// TIA Portal project "Three_Pump_Booster_Control" (V19)
// Three-pump VFD booster station with PID pressure control, lead/lag sequencing and WinCC HMI

(* hardware
DEVICE "S7-1500/ET200MP station_1"  S7-1500 station
   slot 0: "Rail_0"  Rack  6ES7 590-1***0-0AA0
   slot 1: "PLC_Booster"  CPU 1511-1 PN  6ES7 511-1AK02-0AB0  V2.9
      slot 3: "CPU display_1"  6ES7591-1AA00-0AA0
      slot 32768: "PROFINET interface_1"  X1
         slot 32769: "Port_1"  X1 P1
         slot 32770: "Port_2"  X1 P2
      slot 34817: "Virtual CP interface port_1"  Virtual CP interface port  Virtual CP interface port
DEVICE "HMI_Booster"  SIMATIC PC station
   slot 0: "SIMATIC PC station"  Rail  SIMATIC PC-Station  V1.0
      slot 125: "Stationmanager"  Station_Manager  V6.0.4
   slot 1: "HMI_RT_1"  WinCC RT Advanced  6AV2 104-0xxxx-xxxx  17.0.0.0
      slot 33792: "Computer interface"  Host interface
   slot 2: "IE general_1"  IE General  IE_CP  V8.2.0
      slot 1: "PROFINET interface"  IEGeneral.Interface.8.2.0
*)

// ===== PLC "PLC_Booster"  CPU 1511-1 PN =====

TYPE "UDT_Pump"
   STRUCT
      CmdRun : Bool;
      CmdSpeedPct : Real;
      FbRunning : Bool;
      FbFault : Bool;
      FbSpeedPct : Real;
      RunHours : Real;
      Role : Int;
   END_STRUCT;
END_TYPE

DATA_BLOCK "DB_Pumps"   // DB1
{ S7_Optimized_Access := 'TRUE' }
VERSION : 0.1
   VAR
      Pump1 : "UDT_Pump";
      Pump2 : "UDT_Pump";
      Pump3 : "UDT_Pump";
   END_VAR
BEGIN
END_DATA_BLOCK

DATA_BLOCK "DB_System"   // DB2
{ S7_Optimized_Access := 'TRUE' }
VERSION : 0.1
   VAR
      SystemRun : Bool;
      AutoMode : Bool := TRUE;
      SimEnable : Bool := TRUE;
      PressureSP : Real := 4.0;
      PressurePV : Real;
      PIDOutputPct : Real;
      DemandPct : Real := 35.0;
      PressureHighSP : Real := 6.0;
      PressureLowSP : Real := 2.0;
      PIDMode : Int := 4;
      PIDModeActivate : Bool;
      Pump1RunReq : Bool;
      Pump2RunReq : Bool;
      Pump3RunReq : Bool;
      Pump1SpeedReq : Real;
      Pump2SpeedReq : Real;
      Pump3SpeedReq : Real;
      PumpPermissive : Bool := TRUE;
      Pump1FaultAlarm : Bool;
      Pump2FaultAlarm : Bool;
      Pump3FaultAlarm : Bool;
      PressureHighAlarm : Bool;
      PressureLowAlarm : Bool;
      AnyAlarm : Bool;
      Pump1Role : Int;
      Pump2Role : Int;
      Pump3Role : Int;
      AlarmWord : Word := W#16#0000;
   END_VAR
BEGIN
END_DATA_BLOCK

DATA_BLOCK "DB_Pump1_Control"   // DB3
{ S7_Optimized_Access := 'TRUE' }
VERSION : 0.1
// stored: InstanceOfName FB_PumpControl
"FB_PumpControl"
BEGIN
END_DATA_BLOCK

DATA_BLOCK "DB_Pump2_Control"   // DB4
{ S7_Optimized_Access := 'TRUE' }
VERSION : 0.1
// stored: InstanceOfName FB_PumpControl
"FB_PumpControl"
BEGIN
END_DATA_BLOCK

DATA_BLOCK "DB_Pump3_Control"   // DB5
{ S7_Optimized_Access := 'TRUE' }
VERSION : 0.1
// stored: InstanceOfName FB_PumpControl
"FB_PumpControl"
BEGIN
END_DATA_BLOCK

DATA_BLOCK "DB_ProcessSimulation"   // DB6
{ S7_Optimized_Access := 'TRUE' }
VERSION : 0.1
// stored: InstanceOfName FB_ProcessSimulation
"FB_ProcessSimulation"
BEGIN
END_DATA_BLOCK

DATA_BLOCK "DB_PumpManager"   // DB8
{ S7_Optimized_Access := 'TRUE' }
VERSION : 0.1
// stored: InstanceOfName FB_PumpManager
"FB_PumpManager"
BEGIN
END_DATA_BLOCK

DATA_BLOCK "DB_AlarmManager"   // DB9
{ S7_Optimized_Access := 'TRUE' }
VERSION : 0.1
// stored: InstanceOfName FB_AlarmManager
"FB_AlarmManager"
BEGIN
END_DATA_BLOCK

FUNCTION_BLOCK "FB_PumpControl"   // FB1, LAD
{ S7_Optimized_Access := 'TRUE' }
VERSION : 0.1
   VAR_INPUT
      RunRequest : Bool;
      SpeedRequestPct : Real;
      Permissive : Bool;
   END_VAR
   VAR_IN_OUT
      Pump : "UDT_Pump";
   END_VAR
   VAR_TEMP
      LimitedSpeedPct : Real;
   END_VAR
BEGIN

REGION Network 1: VFD Run Command
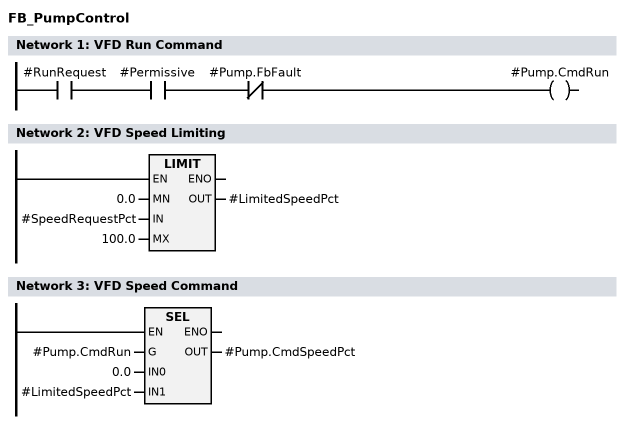
   RUNG wire#powerrail
      Contact( #RunRequest )
      Contact( #Permissive )
      I_Contact( #Pump.FbFault )
      Coil( #Pump.CmdRun )
   END_RUNG
   // the same network as SCL:
   #Pump.CmdRun := #RunRequest AND #Permissive AND NOT #Pump.FbFault;
END_REGION

REGION Network 2: VFD Speed Limiting
   #LimitedSpeedPct := LIMIT(MN := 0.0, IN := #SpeedRequestPct, MX := 100.0);
END_REGION

REGION Network 3: VFD Speed Command
   #Pump.CmdSpeedPct := SEL(G := #Pump.CmdRun, IN0 := 0.0, IN1 := #LimitedSpeedPct);
END_REGION
END_FUNCTION_BLOCK

FUNCTION_BLOCK "FB_ProcessSimulation"   // FB2, SCL
{ S7_Optimized_Access := 'TRUE' }
VERSION : 0.1
   VAR_INPUT
      SimEnable : Bool;
      DemandPct : Real;
   END_VAR
   VAR_IN_OUT
      Pump1 : "UDT_Pump";
      Pump2 : "UDT_Pump";
      Pump3 : "UDT_Pump";
      PressurePV : Real;
   END_VAR
   VAR_TEMP
      TargetSpeed1 : Real;
      TargetSpeed2 : Real;
      TargetSpeed3 : Real;
      TotalFlow : Real;
      DemandLimited : Real;
   END_VAR
BEGIN

   IF NOT #SimEnable THEN
       // Reset simulated process
       #Pump1.FbSpeedPct := 0.0;
       #Pump2.FbSpeedPct := 0.0;
       #Pump3.FbSpeedPct := 0.0;

       #Pump1.FbRunning := FALSE;
       #Pump2.FbRunning := FALSE;
       #Pump3.FbRunning := FALSE;

       #PressurePV := 0.0;

   ELSE
       // Determine requested VFD speeds
       #TargetSpeed1 := 0.0;
       #TargetSpeed2 := 0.0;
       #TargetSpeed3 := 0.0;

       IF #Pump1.CmdRun AND NOT #Pump1.FbFault THEN
           #TargetSpeed1 := #Pump1.CmdSpeedPct;
       END_IF;

       IF #Pump2.CmdRun AND NOT #Pump2.FbFault THEN
           #TargetSpeed2 := #Pump2.CmdSpeedPct;
       END_IF;

       IF #Pump3.CmdRun AND NOT #Pump3.FbFault THEN
           #TargetSpeed3 := #Pump3.CmdSpeedPct;
       END_IF;

       // Simulate VFD acceleration and deceleration
       #Pump1.FbSpeedPct := #Pump1.FbSpeedPct +
       0.2 * (#TargetSpeed1 - #Pump1.FbSpeedPct);

       #Pump2.FbSpeedPct := #Pump2.FbSpeedPct +
       0.2 * (#TargetSpeed2 - #Pump2.FbSpeedPct);

       #Pump3.FbSpeedPct := #Pump3.FbSpeedPct +
       0.2 * (#TargetSpeed3 - #Pump3.FbSpeedPct);

       // Simulated running feedback
       #Pump1.FbRunning := #Pump1.FbSpeedPct > 1.0;
       #Pump2.FbRunning := #Pump2.FbSpeedPct > 1.0;
       #Pump3.FbRunning := #Pump3.FbSpeedPct > 1.0;

       // Combined pump flow (arbitrary simulation units)
       #TotalFlow := 1.1 * (
       #Pump1.FbSpeedPct +
       #Pump2.FbSpeedPct +
       #Pump3.FbSpeedPct
       );

       // Limit simulated water demand
       #DemandLimited := #DemandPct;

       IF #DemandLimited < 0.0 THEN
           #DemandLimited := 0.0;
       ELSIF #DemandLimited > 100.0 THEN
           #DemandLimited := 100.0;
       END_IF;

       // Pressure model: designed for a 100 ms cycle
       #PressurePV := #PressurePV + 0.004 *
       (#TotalFlow - #DemandLimited -
       12.0 * #PressurePV);

       // Limit simulated pressure to 0-10 bar
       IF #PressurePV < 0.0 THEN
           #PressurePV := 0.0;
       ELSIF #PressurePV > 10.0 THEN
           #PressurePV := 10.0;
       END_IF;

   END_IF;
END_FUNCTION_BLOCK

FUNCTION_BLOCK "FB_PumpManager"   // FB3, SCL
{ S7_Optimized_Access := 'TRUE' }
VERSION : 0.1
   VAR_INPUT
      SystemRun : Bool;
      AutoMode : Bool;
      SimEnable : Bool;
      PumpPermissive : Bool;
      PressureSP : Real;
      PressurePV : Real;
      PIDOutputPct : Real;
      Pump1Fault : Bool;
      Pump2Fault : Bool;
      Pump3Fault : Bool;
   END_VAR
   VAR_OUTPUT
      Pump1RunReq : Bool;
      Pump2RunReq : Bool;
      Pump3RunReq : Bool;
      Pump1SpeedReq : Real;
      Pump2SpeedReq : Real;
      Pump3SpeedReq : Real;
      Pump1Role : Int;
      Pump2Role : Int;
      Pump3Role : Int;
   END_VAR
   VAR
      LagActive : Bool;
      StageUpCount : Int := 0;
      StageDownCount : Int;
      LeadPumpNo : Int := 1;
      LagPumpNo : Int;
   END_VAR
   VAR_TEMP
      PreviousLead : Int;
   END_VAR
BEGIN

   (* Default pump commands *)
   #Pump1RunReq := FALSE;
   #Pump2RunReq := FALSE;
   #Pump3RunReq := FALSE;

   #Pump1SpeedReq := 0.0;
   #Pump2SpeedReq := 0.0;
   #Pump3SpeedReq := 0.0;

   IF NOT (#SystemRun AND #AutoMode AND
       #SimEnable AND #PumpPermissive) THEN

       // Reset assignments when system stops
       #LeadPumpNo := 1;
       #LagPumpNo := 0;
       #LagActive := FALSE;
       #StageUpCount := 0;
       #StageDownCount := 0;

   ELSE

       #PreviousLead := #LeadPumpNo;

       // Check the selected lead pump
       CASE #LeadPumpNo OF

           1:
               IF #Pump1Fault THEN
                   IF NOT #Pump3Fault THEN
                       #LeadPumpNo := 3;
                   ELSIF NOT #Pump2Fault THEN
                       #LeadPumpNo := 2;
                   ELSE
                       #LeadPumpNo := 0;
                   END_IF;
               END_IF;

           2:
               IF #Pump2Fault THEN
                   IF NOT #Pump3Fault THEN
                       #LeadPumpNo := 3;
                   ELSIF NOT #Pump1Fault THEN
                       #LeadPumpNo := 1;
                   ELSE
                       #LeadPumpNo := 0;
                   END_IF;
               END_IF;

           3:
               IF #Pump3Fault THEN
                   IF NOT #Pump2Fault THEN
                       #LeadPumpNo := 2;
                   ELSIF NOT #Pump1Fault THEN
                       #LeadPumpNo := 1;
                   ELSE
                       #LeadPumpNo := 0;
                   END_IF;
               END_IF;

           ELSE
               // Recover when a pump becomes available
               IF NOT #Pump1Fault THEN
                   #LeadPumpNo := 1;
               ELSIF NOT #Pump3Fault THEN
                   #LeadPumpNo := 3;
               ELSIF NOT #Pump2Fault THEN
                   #LeadPumpNo := 2;
               ELSE
                   #LeadPumpNo := 0;
               END_IF;

       END_CASE;

       // Reset staging after lead changeover
       IF #LeadPumpNo <> #PreviousLead THEN
           #LagActive := FALSE;
           #LagPumpNo := 0;
           #StageUpCount := 0;
           #StageDownCount := 0;
       END_IF;

       // Check an active assist pump for faults
       IF #LagActive THEN

           IF ((#LagPumpNo = 1) AND #Pump1Fault) OR
               ((#LagPumpNo = 2) AND #Pump2Fault) OR
               ((#LagPumpNo = 3) AND #Pump3Fault) OR
               (#LagPumpNo = #LeadPumpNo) THEN

               #LagPumpNo := 0;

               // Select another healthy assist pump
               CASE #LeadPumpNo OF

                   1:
                       IF NOT #Pump2Fault THEN
                           #LagPumpNo := 2;
                       ELSIF NOT #Pump3Fault THEN
                           #LagPumpNo := 3;
                       END_IF;

                   2:
                       IF NOT #Pump3Fault THEN
                           #LagPumpNo := 3;
                       ELSIF NOT #Pump1Fault THEN
                           #LagPumpNo := 1;
                       END_IF;

                   3:
                       IF NOT #Pump2Fault THEN
                           #LagPumpNo := 2;
                       ELSIF NOT #Pump1Fault THEN
                           #LagPumpNo := 1;
                       END_IF;

               END_CASE;

               IF #LagPumpNo = 0 THEN
                   #LagActive := FALSE;
               END_IF;

           END_IF;

       END_IF;

       // Automatic lag pump staging
       IF NOT #LagActive THEN

           #StageDownCount := 0;

           IF (#LeadPumpNo <> 0) AND
               (#PIDOutputPct >= 95.0) AND
               (#PressurePV < (#PressureSP - 0.2)) THEN

               IF #StageUpCount < 50 THEN
                   #StageUpCount := #StageUpCount + 1;
               END_IF;

           ELSE
               #StageUpCount := 0;
           END_IF;

           IF #StageUpCount >= 50 THEN

               #LagPumpNo := 0;

               CASE #LeadPumpNo OF

                   1:
                       IF NOT #Pump2Fault THEN
                           #LagPumpNo := 2;
                       ELSIF NOT #Pump3Fault THEN
                           #LagPumpNo := 3;
                       END_IF;

                   2:
                       IF NOT #Pump3Fault THEN
                           #LagPumpNo := 3;
                       ELSIF NOT #Pump1Fault THEN
                           #LagPumpNo := 1;
                       END_IF;

                   3:
                       IF NOT #Pump2Fault THEN
                           #LagPumpNo := 2;
                       ELSIF NOT #Pump1Fault THEN
                           #LagPumpNo := 1;
                       END_IF;

               END_CASE;

               #LagActive := (#LagPumpNo <> 0);
               #StageUpCount := 0;

           END_IF;

       ELSE

           #StageUpCount := 0;

           IF (#PIDOutputPct <= 50.0) AND
               (#PressurePV >= (#PressureSP - 0.1)) THEN

               IF #StageDownCount < 100 THEN
                   #StageDownCount := #StageDownCount + 1;
               END_IF;

           ELSE
               #StageDownCount := 0;
           END_IF;

           IF #StageDownCount >= 100 THEN
               #LagActive := FALSE;
               #LagPumpNo := 0;
               #StageDownCount := 0;
           END_IF;

       END_IF;

       // Assign PID speed to selected lead pump
       CASE #LeadPumpNo OF

           1:
               #Pump1RunReq := TRUE;
               #Pump1SpeedReq := #PIDOutputPct;

           2:
               #Pump2RunReq := TRUE;
               #Pump2SpeedReq := #PIDOutputPct;

           3:
               #Pump3RunReq := TRUE;
               #Pump3SpeedReq := #PIDOutputPct;

       END_CASE;

       // Assign fixed 30% speed to assist pump
       IF #LagActive THEN

           CASE #LagPumpNo OF

               1:
                   #Pump1RunReq := TRUE;
                   #Pump1SpeedReq := 30.0;

               2:
                   #Pump2RunReq := TRUE;
                   #Pump2SpeedReq := 30.0;

               3:
                   #Pump3RunReq := TRUE;
                   #Pump3SpeedReq := 30.0;

           END_CASE;

       END_IF;

   END_IF;


   // Default: All pumps on standby
   #Pump1Role := 0;
   #Pump2Role := 0;
   #Pump3Role := 0;

   // Assign operating roles when system enabled
   IF #SystemRun AND #AutoMode AND
       #SimEnable AND #PumpPermissive THEN

       // Lead pump role
       CASE #LeadPumpNo OF
           1:
               #Pump1Role := 1;
           2:
               #Pump2Role := 1;
           3:
               #Pump3Role := 1;
       END_CASE;

       // Assist pump role
       IF #LagActive THEN
           CASE #LagPumpNo OF
               1:
                   #Pump1Role := 2;
               2:
                   #Pump2Role := 2;
               3:
                   #Pump3Role := 2;
           END_CASE;
       END_IF;

   END_IF;

   // Fault indication takes priority
   IF #Pump1Fault THEN
       #Pump1Role := 3;
   END_IF;

   IF #Pump2Fault THEN
       #Pump2Role := 3;
   END_IF;

   IF #Pump3Fault THEN
       #Pump3Role := 3;
   END_IF;
END_FUNCTION_BLOCK

FUNCTION_BLOCK "FB_AlarmManager"   // FB4, SCL
{ S7_Optimized_Access := 'TRUE' }
VERSION : 0.1
   VAR_INPUT
      SystemRun : Bool;
      PressurePV : Real;
      PressureHighSP : Real;
      PressureLowSP : Real;
      Pump1Fault : Bool;
      Pump2Fault : Bool;
      Pump3Fault : Bool;
   END_VAR
   VAR_OUTPUT
      Pump1FaultAlarm : Bool;
      Pump2FaultAlarm : Bool;
      Pump3FaultAlarm : Bool;
      PressureHighAlarm : Bool;
      PressureLowAlarm : Bool;
      AnyAlarm : Bool;
      AlarmWord : Word;
   END_VAR
   VAR
      LowPressureCount : Int;
   END_VAR
BEGIN

   // Individual pump fault alarms
   #Pump1FaultAlarm := #Pump1Fault;
   #Pump2FaultAlarm := #Pump2Fault;
   #Pump3FaultAlarm := #Pump3Fault;

   // High pressure alarm with hysteresis
   IF #PressurePV >= #PressureHighSP THEN
       #PressureHighAlarm := TRUE;
   ELSIF #PressurePV <= (#PressureHighSP - 0.2) THEN
       #PressureHighAlarm := FALSE;
   END_IF;

   // Low pressure alarm with 10-second delay
   // FB must execute every 100 ms
   IF NOT #SystemRun THEN
       #LowPressureCount := 0;
       #PressureLowAlarm := FALSE;

   ELSIF #PressurePV < #PressureLowSP THEN
       IF #LowPressureCount < 100 THEN
           #LowPressureCount := #LowPressureCount + 1;
       END_IF;

       IF #LowPressureCount >= 100 THEN
           #PressureLowAlarm := TRUE;
       END_IF;

   ELSE
       #LowPressureCount := 0;

       IF #PressurePV >= (#PressureLowSP + 0.2) THEN
           #PressureLowAlarm := FALSE;
       END_IF;
   END_IF;

   // General alarm indication
   #AnyAlarm :=
   #Pump1FaultAlarm OR
   #Pump2FaultAlarm OR
   #Pump3FaultAlarm OR
   #PressureHighAlarm OR
   #PressureLowAlarm;



   // Pack individual alarm signals
   // into one WinCC alarm trigger word

   #AlarmWord := W#16#0000;

   IF #Pump1FaultAlarm THEN
       #AlarmWord := #AlarmWord OR W#16#0001;
   END_IF;

   IF #Pump2FaultAlarm THEN
       #AlarmWord := #AlarmWord OR W#16#0002;
   END_IF;

   IF #Pump3FaultAlarm THEN
       #AlarmWord := #AlarmWord OR W#16#0004;
   END_IF;

   IF #PressureHighAlarm THEN
       #AlarmWord := #AlarmWord OR W#16#0008;
   END_IF;

   IF #PressureLowAlarm THEN
       #AlarmWord := #AlarmWord OR W#16#0010;
   END_IF;
END_FUNCTION_BLOCK

ORGANIZATION_BLOCK "Main"   // OB1, LAD, ProgramCycle
TITLE = "Main Program Sweep (Cycle)"
{ S7_Optimized_Access := 'TRUE' }
VERSION : 0.1
   VAR_INPUT
      Initial_Call : Bool;   // Initial call of this OB
      Remanence : Bool;   // =True, if remanent data are available
   END_VAR
BEGIN

REGION Network 1: Pump 1 VFD Control
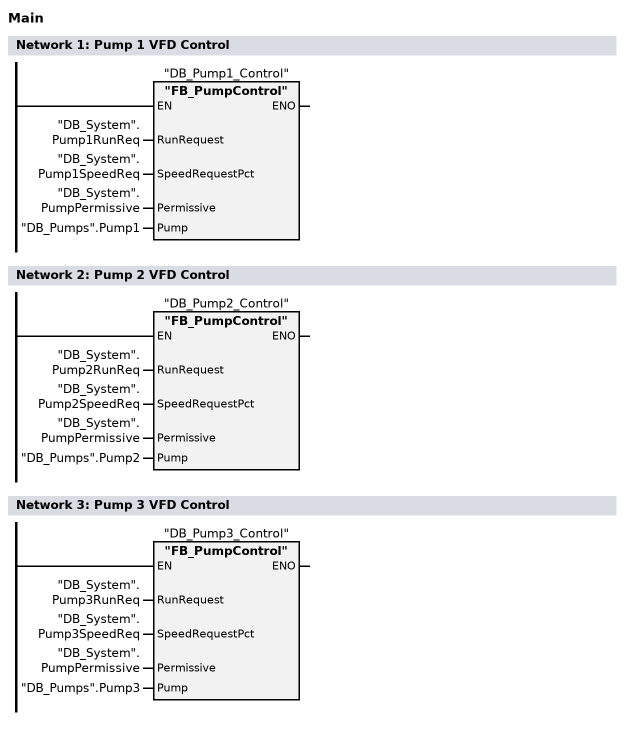
   RUNG wire#powerrail
      "DB_Pump1_Control"(RunRequest := "DB_System".Pump1RunReq, SpeedRequestPct := "DB_System".Pump1SpeedReq, Permissive := "DB_System".PumpPermissive, Pump := "DB_Pumps".Pump1)
   END_RUNG
   // the same network as SCL:
   "DB_Pump1_Control"(RunRequest := "DB_System".Pump1RunReq,   // "FB_PumpControl"
                      SpeedRequestPct := "DB_System".Pump1SpeedReq,
                      Permissive := "DB_System".PumpPermissive,
                      Pump := "DB_Pumps".Pump1);
END_REGION

REGION Network 2: Pump 2 VFD Control
   RUNG wire#powerrail
      "DB_Pump2_Control"(RunRequest := "DB_System".Pump2RunReq, SpeedRequestPct := "DB_System".Pump2SpeedReq, Permissive := "DB_System".PumpPermissive, Pump := "DB_Pumps".Pump2)
   END_RUNG
   // the same network as SCL:
   "DB_Pump2_Control"(RunRequest := "DB_System".Pump2RunReq,   // "FB_PumpControl"
                      SpeedRequestPct := "DB_System".Pump2SpeedReq,
                      Permissive := "DB_System".PumpPermissive,
                      Pump := "DB_Pumps".Pump2);
END_REGION

REGION Network 3: Pump 3 VFD Control
   RUNG wire#powerrail
      "DB_Pump3_Control"(RunRequest := "DB_System".Pump3RunReq, SpeedRequestPct := "DB_System".Pump3SpeedReq, Permissive := "DB_System".PumpPermissive, Pump := "DB_Pumps".Pump3)
   END_RUNG
   // the same network as SCL:
   "DB_Pump3_Control"(RunRequest := "DB_System".Pump3RunReq,   // "FB_PumpControl"
                      SpeedRequestPct := "DB_System".Pump3SpeedReq,
                      Permissive := "DB_System".PumpPermissive,
                      Pump := "DB_Pumps".Pump3);
END_REGION
END_ORGANIZATION_BLOCK

ORGANIZATION_BLOCK "OB30_ProcessControl"   // OB30, LAD, CyclicInterrupt
{ S7_Optimized_Access := 'TRUE' }
VERSION : 0.1
   VAR_INPUT
      Initial_Call : Bool;   // Initial call of this OB
      Event_Count : Int;   // Events discarded
   END_VAR
BEGIN

REGION Network 1: Hydraulic Process Simulation
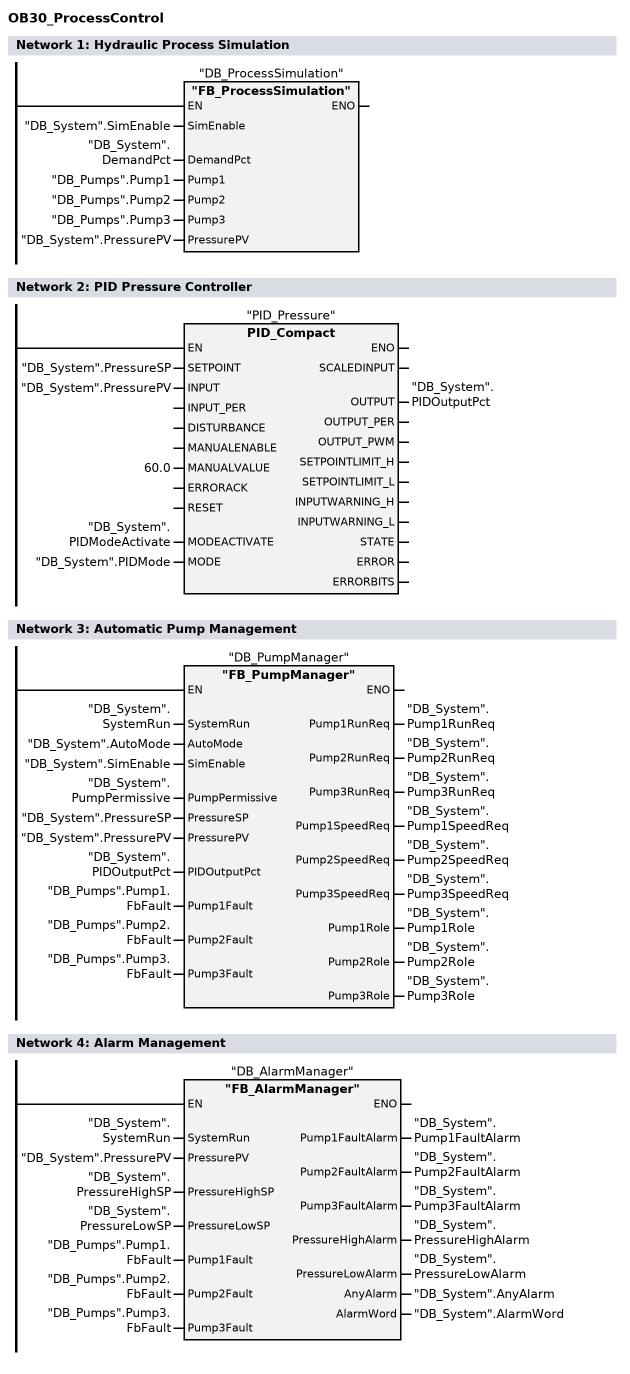
   RUNG wire#powerrail
      "DB_ProcessSimulation"(SimEnable := "DB_System".SimEnable, DemandPct := "DB_System".DemandPct, Pump1 := "DB_Pumps".Pump1, Pump2 := "DB_Pumps".Pump2, Pump3 := "DB_Pumps".Pump3, PressurePV := "DB_System".PressurePV)
   END_RUNG
   // the same network as SCL:
   "DB_ProcessSimulation"(SimEnable := "DB_System".SimEnable,   // "FB_ProcessSimulation"
                          DemandPct := "DB_System".DemandPct,
                          Pump1 := "DB_Pumps".Pump1,
                          Pump2 := "DB_Pumps".Pump2,
                          Pump3 := "DB_Pumps".Pump3,
                          PressurePV := "DB_System".PressurePV);
END_REGION

REGION Network 2: PID Pressure Controller
   "PID_Pressure"(Setpoint := "DB_System".PressureSP,   // PID_Compact
                  Input := "DB_System".PressurePV,
                  ManualValue := 60.0,
                  ModeActivate := "DB_System".PIDModeActivate,
                  Mode := "DB_System".PIDMode,
                  Output => "DB_System".PIDOutputPct);
END_REGION

REGION Network 3: Automatic Pump Management
   RUNG wire#powerrail
      "DB_PumpManager"(SystemRun := "DB_System".SystemRun, AutoMode := "DB_System".AutoMode, SimEnable := "DB_System".SimEnable, PumpPermissive := "DB_System".PumpPermissive, PressureSP := "DB_System".PressureSP, PressurePV := "DB_System".PressurePV, PIDOutputPct := "DB_System".PIDOutputPct, Pump1Fault := "DB_Pumps".Pump1.FbFault, Pump2Fault := "DB_Pumps".Pump2.FbFault, Pump3Fault := "DB_Pumps".Pump3.FbFault, Pump1RunReq => "DB_System".Pump1RunReq, Pump2RunReq => "DB_System".Pump2RunReq, Pump3RunReq => "DB_System".Pump3RunReq, Pump1SpeedReq => "DB_System".Pump1SpeedReq, Pump2SpeedReq => "DB_System".Pump2SpeedReq, Pump3SpeedReq => "DB_System".Pump3SpeedReq, Pump1Role => "DB_System".Pump1Role, Pump2Role => "DB_System".Pump2Role, Pump3Role => "DB_System".Pump3Role)
   END_RUNG
   // the same network as SCL:
   "DB_PumpManager"(SystemRun := "DB_System".SystemRun,   // "FB_PumpManager"
                    AutoMode := "DB_System".AutoMode,
                    SimEnable := "DB_System".SimEnable,
                    PumpPermissive := "DB_System".PumpPermissive,
                    PressureSP := "DB_System".PressureSP,
                    PressurePV := "DB_System".PressurePV,
                    PIDOutputPct := "DB_System".PIDOutputPct,
                    Pump1Fault := "DB_Pumps".Pump1.FbFault,
                    Pump2Fault := "DB_Pumps".Pump2.FbFault,
                    Pump3Fault := "DB_Pumps".Pump3.FbFault,
                    Pump1RunReq => "DB_System".Pump1RunReq,
                    Pump2RunReq => "DB_System".Pump2RunReq,
                    Pump3RunReq => "DB_System".Pump3RunReq,
                    Pump1SpeedReq => "DB_System".Pump1SpeedReq,
                    Pump2SpeedReq => "DB_System".Pump2SpeedReq,
                    Pump3SpeedReq => "DB_System".Pump3SpeedReq,
                    Pump1Role => "DB_System".Pump1Role,
                    Pump2Role => "DB_System".Pump2Role,
                    Pump3Role => "DB_System".Pump3Role);
END_REGION

REGION Network 4: Alarm Management
   RUNG wire#powerrail
      "DB_AlarmManager"(SystemRun := "DB_System".SystemRun, PressurePV := "DB_System".PressurePV, PressureHighSP := "DB_System".PressureHighSP, PressureLowSP := "DB_System".PressureLowSP, Pump1Fault := "DB_Pumps".Pump1.FbFault, Pump2Fault := "DB_Pumps".Pump2.FbFault, Pump3Fault := "DB_Pumps".Pump3.FbFault, Pump1FaultAlarm => "DB_System".Pump1FaultAlarm, Pump2FaultAlarm => "DB_System".Pump2FaultAlarm, Pump3FaultAlarm => "DB_System".Pump3FaultAlarm, PressureHighAlarm => "DB_System".PressureHighAlarm, PressureLowAlarm => "DB_System".PressureLowAlarm, AnyAlarm => "DB_System".AnyAlarm, AlarmWord => "DB_System".AlarmWord)
   END_RUNG
   // the same network as SCL:
   "DB_AlarmManager"(SystemRun := "DB_System".SystemRun,   // "FB_AlarmManager"
                     PressurePV := "DB_System".PressurePV,
                     PressureHighSP := "DB_System".PressureHighSP,
                     PressureLowSP := "DB_System".PressureLowSP,
                     Pump1Fault := "DB_Pumps".Pump1.FbFault,
                     Pump2Fault := "DB_Pumps".Pump2.FbFault,
                     Pump3Fault := "DB_Pumps".Pump3.FbFault,
                     Pump1FaultAlarm => "DB_System".Pump1FaultAlarm,
                     Pump2FaultAlarm => "DB_System".Pump2FaultAlarm,
                     Pump3FaultAlarm => "DB_System".Pump3FaultAlarm,
                     PressureHighAlarm => "DB_System".PressureHighAlarm,
                     PressureLowAlarm => "DB_System".PressureLowAlarm,
                     AnyAlarm => "DB_System".AnyAlarm,
                     AlarmWord => "DB_System".AlarmWord);
END_REGION
END_ORGANIZATION_BLOCK

(* ===== HMI "HMI_RT_1" =====
system functions are stored by id; their names below are inferred from use
connection "HMI_Connection_1": ETHERNET, S7_1500_OMS

HMI tags "Default tag table"
   "HMI_PressurePV" : Real = PLC DB_System.PressurePV AT %DB1.DBD0, 1 s
   "HMI_PressureSP" : Real = PLC DB_System.PressureSP AT %DB1.DBD0, 1 s
   "HMI_TestValue" : Real AT %DB1.DBD0
   "HMI_P1_Running" : Bool = PLC DB_Pumps.Pump1.FbRunning AT %DB1.DBX0.0, 1 s
   "HMI_P2_Running" : Bool = PLC DB_Pumps.Pump2.FbRunning AT %DB1.DBX0.0, 1 s
   "HMI_P3_Running" : Bool = PLC DB_Pumps.Pump3.FbRunning AT %DB1.DBX0.0, 1 s
   "HMI_P1_Speed" : Real = PLC DB_Pumps.Pump1.FbSpeedPct AT %DB1.DBX0.0, 1 s
   "HMI_P2_Speed" : Real = PLC DB_Pumps.Pump2.FbSpeedPct AT %DB1.DBD0, 1 s
   "HMI_P3_Speed" : Real = PLC DB_Pumps.Pump3.FbSpeedPct AT %DB1.DBD0, 1 s
   "HMI_SystemRun" : Bool = PLC DB_System.SystemRun AT %DB1.DBX0.0, 1 s
   "HMI_PIDOutput" : Real = PLC DB_System.PIDOutputPct AT %DB1.DBD0, 1 s
   "HMI_P1_Role" : Int = PLC DB_System.Pump1Role AT %DB1.DBW0, 1 s
   "HMI_P2_Role" : Int = PLC DB_System.Pump2Role AT %DB1.DBW0, 1 s
   "HMI_P3_Role" : Int = PLC DB_System.Pump3Role AT %DB1.DBW0, 1 s
   "HMI_DemandPct" : Real = PLC DB_System.DemandPct AT %DB1.DBD0, 1 s
   "HMI_AutoMode" : Bool = PLC DB_System.AutoMode AT %DB1.DBX0.0, 1 s
   "HMI_AnyAlarm" : Bool = PLC DB_System.AnyAlarm AT %DB1.DBX0.0, 1 s
   "PID_ACTIVE" : Bool = PLC DB_System.PIDModeActivate AT %DB1.DBX0.0, 1 s
   "HMI_AlarmWord" : Word = PLC DB_System.AlarmWord AT %DB1.DBW0, 1 s
   "PID_DeActive" : Bool = PLC DB_System.PIDModeActivate AT %DB1.DBX0.0, 1 s
      on ChangeValue: ResetBit("PID_DeActive")

discrete alarms
   1: 'PUMP 01 - VFD FAULT', class Errors, trigger "HMI_AlarmWord" bit 0
   2: 'PUMP 02 - VFD FAULT', class Errors, trigger "HMI_AlarmWord" bit 1
   3: 'PUMP 03 - VFD FAULT', class Errors, trigger "HMI_AlarmWord" bit 2
   4: 'HIGH DISCHARGE PRESSURE', class Warnings, trigger "HMI_AlarmWord" bit 3
   5: 'LOW DISCHARGE PRESSURE', class Warnings, trigger "HMI_AlarmWord" bit 4

text list "TL_PumpRole": 0 'STANDBY'; 1 'LEAD'; 2 'ASSIST'; 3 'FAULT'

text list "TL_SystemStatus": 0 'STOPPED'; 1 'ENABLED'

text list "TL_OperatingMode": 0 'MANUAL'; 1 'AUTO'

text list "TL_AlarmStatus": 0 'NO ACTIVE ALARMS'; 1 'ALARM ACTIVE'

screen "01_Overview" 1024x768
   TextField "Text field_12" at 28,232 size 241x22; Text 'PUMP STATUS & VFD CONTROL'
   IOField "I/O field_1" at 48,150 size 90x32; FormatPattern 9.99
      ProcessValue <- "HMI_PressurePV"
   TextField "Text field_1" at 48,115 size 180x22; Text 'DISCHARGE PRESSURE'
   IOField "I/O field_2" at 379,150 size 79x32; FormatPattern 9.99
      ProcessValue <- "HMI_PressureSP"
   TextField "Text field_2" at 379,115 size 168x22; Text 'PRESSURE SETPOINT'
   Circle "Circle_1" at 294,285 size 20x20
      Appearance <- "HMI_P1_Running"
   TextField "Text field_3" at 48,285 size 73x22; Text 'PUMP 01'
   IOField "I/O field_3" at 143,330 size 75x32; FormatPattern 99.9
      ProcessValue <- "HMI_P1_Speed"
   TextField "Text field_4" at 125,377 size 124x22; Text 'VFD SPEED (%)'
   Circle "Circle_2" at 617,285 size 20x20
      Appearance <- "HMI_P2_Running"
   TextField "Text field_5" at 379,285 size 73x22; Text 'PUMP 02'
   IOField "I/O field_4" at 468,330 size 69x32; FormatPattern 99.9
      ProcessValue <- "HMI_P2_Speed"
   TextField "Text field_6" at 436,373 size 124x22; Text 'VFD SPEED (%)'
   Circle "Circle_3" at 947,285 size 20x20
      Appearance <- "HMI_P3_Running"
   TextField "Text field_7" at 710,285 size 73x22; Text 'PUMP 03'
   IOField "I/O field_5" at 805,330 size 76x32; FormatPattern 99.9
      ProcessValue <- "HMI_P3_Speed"
   TextField "Text field_8" at 793,373 size 124x22; Text 'VFD SPEED (%)'
   Button "Button_1" at 43,566 size 125x46; TextOff 'START SYSTEM'
      on Press: SetBit("HMI_SystemRun")
   Button "Button_2" at 190,566 size 120x46; TextOff 'STOP SYSTEM'
      on Press: ResetBit("HMI_SystemRun")
   Circle "Circle_4" at 713,566 size 22x22
      Appearance <- "HMI_SystemRun"
   TextField "Text field_10" at 32,14 size 379x36; Text 'THREE-PUMP BOOSTER STATION'
   TextField "Text field_11" at 34,51 size 232x19; Text 'AUTOMATIC PRESSURE CONTROL SYSTEM'
   TextField "Text field_13" at 48,526 size 146x22; Text 'SYSTEM CONTROL'
   TextField "Text field_14" at 710,526 size 130x22; Text 'SYSTEM STATUS'
   Button "Button_3" at 690,682 size 145x50; TextOff 'TRENDS'
      on Click: ActivateScreen("02_Trends", 0)
   Button "Button_4" at 851,682 size 145x50; TextOff 'ALARMS'
      on Click: ActivateScreen("03_Alarms", 0)
   TextField "Text field_9" at 385,526 size 129x22; Text 'WATER DEMAND'
   Bar "Bar_1" at 48,428 size 266x24; MinimumValue 0; MaximumValue 100
      ProcessValue <- "HMI_P1_Speed"
   TextField "Text field_15" at 48,451 size 22x17; Text '0%'
   TextField "Text field_16" at 158,451 size 28x17; Text '50%'
   TextField "Text field_17" at 268,451 size 34x17; Text '100%'
   Bar "Bar_2" at 378,428 size 266x24; MinimumValue 0; MaximumValue 100
      ProcessValue <- "HMI_P2_Speed"
   TextField "Text field_18" at 378,451 size 22x17; Text '0%'
   TextField "Text field_19" at 488,451 size 28x17; Text '50%'
   TextField "Text field_20" at 598,451 size 34x17; Text '100%'
   Bar "Bar_3" at 708,428 size 266x24; MinimumValue 0; MaximumValue 100
      ProcessValue <- "HMI_P3_Speed"
   TextField "Text field_21" at 708,451 size 22x17; Text '0%'
   TextField "Text field_22" at 818,451 size 28x17; Text '50%'
   TextField "Text field_23" at 928,451 size 34x17; Text '100%'
   TextField "Text field_24" at 710,115 size 99x22; Text 'PID OUTPUT'
   IOField "I/O field_6" at 711,141 size 168x44; FormatPattern 99.9
      ProcessValue <- "HMI_PIDOutput"
   TextField "Text field_25" at 793,149 size 25x25; Text '%'
   TextField "Text field_26" at 463,153 size 33x25; Text 'bar'
   TextField "Text field_27" at 126,153 size 33x25; Text 'bar'
   SymbolicIOField "Symbolic I/O field_1" at 48,399 size 120x20; TextOff '0'; TextOn '1'; TextList "TL_PumpRole"
      ProcessValue <- "HMI_P1_Role"
      Appearance <- "HMI_P1_Role"
   SymbolicIOField "Symbolic I/O field_2" at 379,399 size 120x20; TextOff '0'; TextOn '1'; TextList "TL_PumpRole"
      Appearance <- "HMI_P2_Role"
      ProcessValue <- "HMI_P2_Role"
   SymbolicIOField "Symbolic I/O field_3" at 710,399 size 120x20; TextOff '0'; TextOn '1'; TextList "TL_PumpRole"
      ProcessValue <- "HMI_P3_Role"
      Appearance <- "HMI_P3_Role"
   IOField "I/O field_7" at 379,570 size 125x42; FormatPattern 99.99
      ProcessValue <- "HMI_DemandPct"
   TextField "Text field_28" at 515,577 size 25x25; Text '%'
   TextField "Text field_29" at 376,617 size 204x18; Text 'SIMULATED WATER CONSUMPTION'
   SymbolicIOField "Symbolic I/O field_4" at 750,565 size 205x28; TextOff '0'; TextOn '1'; TextList "TL_SystemStatus"
      ProcessValue <- "HMI_SystemRun"
      Appearance <- "HMI_SystemRun"
   SymbolicIOField "Symbolic I/O field_5" at 865,604 size 105x28; TextOff '0'; TextOn '1'; TextList "TL_OperatingMode"
      ProcessValue <- "HMI_AutoMode"
      Appearance <- "HMI_AutoMode"
   TextField "Text field_30" at 710,607 size 137x21; Text 'OPERATING MODE'
   TextField "Text field_31" at 48,685 size 121x22; Text 'ALARM STATUS'
   Circle "Circle_5" at 226,699 size 18x18
      Appearance <- "HMI_SystemRun"
   SymbolicIOField "Symbolic I/O field_6" at 260,694 size 350x30; TextOff '0'; TextOn '1'; TextList "TL_AlarmStatus"
      Appearance <- "HMI_SystemRun"
      ProcessValue <- "HMI_AnyAlarm"
   Button "Button_5" at 905,141 size 65x32; TextOff 'PID ON'
      on Click: SetBit("PID_ACTIVE")

screen "02_Trends" 1024x768
   TextField "Text field_1" at 32,14 size 363x33; Text 'PRESSURE CONTROL TRENDS'
   TextField "Text field_2" at 34,51 size 264x20; Text 'PID PERFORMANCE & DEMAND RESPONSE'
   TrendView "Trend view_1" at 48,150 size 928x465
      ValueAxis1Begin <- "HMI_PressurePV"
      ValueAxis2Begin <- "HMI_PressureSP"
   TextField "Text field_3" at 48,119 size 180x22; Text 'DISCHARGE PRESSURE'
   TextField "Text field_4" at 735,119 size 182x22; Text 'LIVE PID MONITORING'
   Button "Button_1" at 28,682 size 215x48; TextOff 'BACK TO OVERVIEW'
      on Click: ActivateScreen("01_Overview", 0)

screen "03_Alarms" 1024x768
   TextField "Text field_1" at 32,14 size 363x32; Text 'BOOSTER STATION — ALARMS'
   TextField "Text field_2" at 34,51 size 307x20; Text 'PUMP FAULTS & PRESSURE ALARM MONITORING'
   AlarmView "Alarm view_1" at 48,160 size 928x455
   TextField "Text field_3" at 48,122 size 144x22; Text 'PROCESS ALARMS'
   Button "Button_1" at 34,689 size 169x32; TextOff 'BACK TO OVERVIEW'
      on Click: ActivateScreen("01_Overview", 0)
*)